(* IEC 61131-3 sources: plc-workbench/experiments/general_tasks_r6/final_recheck/natural_language_intake, 2 files *)

(* ---- before.st ---- *)
FUNCTION_BLOCK FanHysteresis
VAR_INPUT
    enabled : BOOL;
    temperature : REAL;
END_VAR
VAR_OUTPUT
    fan : BOOL := FALSE;
END_VAR
VAR CONSTANT
    TEMP_ON : REAL := 30.0;
    TEMP_OFF : REAL := 25.0;
END_VAR

IF NOT enabled THEN
    fan := FALSE;
ELSE
    IF temperature >= TEMP_ON THEN
        fan := TRUE;
    ELSIF temperature <= TEMP_OFF THEN
        fan := FALSE;
    END_IF;
END_IF;
END_FUNCTION_BLOCK

(* ---- candidate_final.st ---- *)
FUNCTION_BLOCK FanHysteresis
VAR_INPUT
    enabled : BOOL;
    temperature : REAL;
END_VAR
VAR_OUTPUT
    fan : BOOL := FALSE;
END_VAR
VAR CONSTANT
    TEMP_ON : REAL := 30.0;
    TEMP_OFF : REAL := 25.0;
END_VAR

IF NOT enabled THEN
    fan := FALSE;
ELSE
    IF temperature >= TEMP_ON THEN
        fan := TRUE;
    ELSIF temperature <= TEMP_OFF THEN
        fan := FALSE;
    END_IF;
END_IF;
END_FUNCTION_BLOCK
